// TIA Portal V20 export
// export: Created 2026-10-12T05:42:34.4695906Z, ExportSetting WithDefaults, DisplayName Totally Integrated Automation Portal, DisplayVersion V20, DisplayName TIA Portal Openness, DisplayVersion V20, DisplayName TIA Portal Teamcenter Gateway, DisplayVersion V20, DisplayName TIA Portal Version Control Interface, DisplayVersion V20, DisplayName SINAMICS Startdrive Advanced, DisplayVersion V20 SP1 Update 2, DisplayName SINAMICS Startdrive G110M, G120, G120C, G120D, G120P, G115D, DisplayVersion V20 SP1 Update 2, DisplayName SINAMICS Startdrive G130, G150, S120, S150, SINAMICS MV, G220, S200, S210, DisplayVersion V20 SP1 Update 2, DisplayName STEP 7 Professional, DisplayVersion V20, DisplayName STEP 7 Safety, DisplayVersion V20, DisplayName WinCC Basic/Comfort/Advanced, DisplayVersion V20, DisplayName WinCC Professional, DisplayVersion V20, DisplayName WinCC Unified, DisplayVersion V20
FUNCTION "F_PressDemoScrap" : Bool   // FC166, SCL
{ S7_Optimized_Access := 'TRUE' }
VERSION : 0.1
// stored: AutoNumber true, IsIECCheckEnabled false, SetENOAutomatically false, UDAEnableTagReadback false
   VAR_IN_OUT
      Seq : "FRK_SequenceCtx";
      Cycle : "ST_PressDemoCycle";
      Core : "FRK_Core";
      Unit : "FRK_Unit";
      Status : "ST_ModuleStatus";
      Part : "ST_PartContext";
      AlarmLog : "FRK_AlarmLog";
   END_VAR
   VAR_TEMP
      Written : Bool;
   END_VAR
BEGIN

   IF "FRK_SeqOnce"(Seq := #Seq, Enable := TRUE, Token := #Seq.Step) THEN
       #Written := "FRK_PartProcessed"(Core := #Core, Unit := #Unit, Status := #Status, Part := #Part, AlarmLog := #AlarmLog,
                                       Verdict := 2, Reason := #Cycle.FailureReason);
       IF NOT #Written AND #Unit.CarrierIndex = 0 AND #Unit.Nok < UDINT#4294967295 THEN
           #Unit.Nok := #Unit.Nok + 1;
           #Unit.NokReason := #Cycle.FailureReason;
       END_IF;
       #Cycle.PartDispositioned := TRUE;
       #Cycle.PartInMachine := FALSE;
       #Cycle.CycleCompleted := FALSE;
   END_IF;
   #F_PressDemoScrap := #Core.Exec <> 3;
END_FUNCTION
